Fanuc KAREL source: KD00064.KL

PROGRAM KD00064
%NOLOCKGROUP
VAR
  I: INTEGER
  J: INTEGER
  B: BOOLEAN
  R: REAL
  S: STRING[80]
BEGIN
  CONDITION[1]:
  WHEN DIN[1] = ON DO
    HOLD
  ENDCONDITION
END KD00064
